VAR_GLOBAL
    // Synchronized snapshot — all data from the same DC cycle.
    // Read from Python via single ADS read: GVL_Sync.stSnapshot
    stSnapshot : ST_SyncSnapshot;
END_VAR

(* stored: Version 1.1.0.1, ProductVersion 3.1.4026.18
   GVL GVL_Sync: Id {f87471bf-b393-4a0a-a16a-0c6d0d0014a0} *)
